FUNCTION VC_GetUInt64 : ULINT
// Reads UInt64 (8 byte, little-endian) from Buf[Pos] and advances Pos.
VAR_IN_OUT
    Buf   : ARRAY[*] OF BYTE;
    Pos   : UDINT;
END_VAR
VAR
    nVal : ULINT;
END_VAR

nVal := 0;
VC_GetRaw(Buf := Buf, Pos := Pos, pDst := ADR(nVal), Size := 8);
VC_GetUInt64 := nVal;

END_FUNCTION

(* stored: Version 1.1.0.1, ProductVersion 3.1.4024.12
   POU VC_GetUInt64: Id {bf7f822e-2a69-43dc-a576-6457b8c60899}, SpecialFunc None *)
